(* IEC 61131-3 sources: axsharp/src/sanbox/integration/ix-integration-plc/src/IO, 5 files *)

(* ---- HwIdentifierList.st ---- *)
NAMESPACE axosimple
    TYPE HwIdentifierList : ARRAY[0..15] OF UINT :=
            [
                UINT#32,
                UINT#48,
                UINT#51,
                UINT#54,
                UINT#64,
                UINT#65,
                UINT#66,
                UINT#72,
                UINT#73,
                UINT#74,
                UINT#117,
                UINT#120,
                UINT#121,
                UINT#135,
                UINT#256,
                UINT#257
    ];
END_TYPE
END_NAMESPACE

(* ---- HwIdentifiers.st ---- *)
NAMESPACE axosimple
    TYPE
        HwIdentifiers : UINT
        (
            plc_line_HwID := UINT#32,
            plc_line_plc_line_HwID := UINT#48,
            plc_line_plc_line_Card_reader_writer_1_HwID := UINT#51,
            plc_line_plc_line_CPU_display_1_HwID := UINT#54,
            plc_line_plc_line_PROFINET_interface_1_HwID := UINT#64,
            plc_line_plc_line_PROFINET_interface_1_Port_1_HwID := UINT#65,
            plc_line_plc_line_PROFINET_interface_1_Port_2_HwID := UINT#66,
            plc_line_plc_line_PROFINET_interface_2_HwID := UINT#72,
            plc_line_plc_line_PROFINET_interface_2_Port_3_HwID := UINT#73,
            plc_line_plc_line_PROFINET_interface_2_Port_4_HwID := UINT#74,
            plc_line_plc_line_OPC_UA_1_HwID := UINT#117,
            plc_line_plc_line_PROFINET_interface_GBIT_3_HwID := UINT#120,
            plc_line_plc_line_PROFINET_interface_GBIT_3_Port_5_HwID := UINT#121,
            plc_line_plc_line_Virtual_communication_interface_HwID := UINT#135,
            profinet_plc_line_HwID := UINT#256,
            plc_line_Rail_0_HwID := UINT#257
        );
    END_TYPE
END_NAMESPACE

(* ---- Inputs.st ---- *)
NAMESPACE axosimple
    TYPE
        {S7.extern=ReadWrite}
        {#ix-attr:[Container(Layout.Wrap)]}
        Inputs : STRUCT
            noInputsFoundInTheHwConfig AT %B0:  BYTE;
        END_STRUCT;
    END_TYPE
END_NAMESPACE

(* ---- Outputs.st ---- *)
NAMESPACE axosimple
    TYPE
        {S7.extern=ReadWrite}
        {#ix-attr:[Container(Layout.Wrap)]}
        Outputs : STRUCT
            noOutputsFoundInTheHwConfig AT %B0:  BYTE;
        END_STRUCT;
    END_TYPE
END_NAMESPACE

(* ---- IoStructures.st ---- *)
NAMESPACE axosimple
END_NAMESPACE
